// TIA Portal V21 export
TagTable "Proto tags"
  P_SwOn : Bool  (PLC tag HMI_IF.SwOn, HMI_Connection_1, 100 ms)
  P_SwOn_q : Bool  (PLC tag "HMI_IF".SwOn, HMI_Connection_1, 100 ms)
  P_Cell : USInt  (PLC tag HMI_IF.CellSt0[0], HMI_Connection_1, 100 ms)
